(* IEC 61131-3 sources: PLC-Static-Analysis/modules/plc-rules/src/test/resources/dev/plca/rules/RulesFuzzTestInputs/fuzzRules, 23 files *)

(* ---- PLCA-Q007_compliant.st ---- *)
FUNCTION F_Twice : INT
VAR_INPUT
    n : INT;
END_VAR
F_Twice := F_Plus(n, n);
END_FUNCTION

FUNCTION F_Plus : INT
VAR_INPUT
    a : INT;
    b : INT;
END_VAR
F_Plus := a + b;
END_FUNCTION

(* ---- PLCA-P001_compliant.st ---- *)
VAR_GLOBAL
    gMode : INT;
    gOk : BOOL;
END_VAR

FUNCTION_BLOCK FB_Ok
VAR_INPUT
    bA : BOOL;
    bB : BOOL;
END_VAR
VAR_OUTPUT
    bOut : BOOL;
    nOut : INT;
END_VAR
VAR
    n : INT;
END_VAR
// default, then override in an IF
bOut := FALSE;
IF bA THEN
    bOut := TRUE;
END_IF
// latches
bOut S= bA;
bOut R= bB;
// sequential use: read in between
nOut := 1;
n := nOut * 2;
nOut := n;
// locals are not coils by default
n := 0;
n := 5;
// mutually exclusive branches
IF bA THEN
    gOk := TRUE;
ELSE
    gOk := FALSE;
END_IF
END_FUNCTION_BLOCK

PROGRAM P_Ok
VAR
    fb : FB_Ok;
END_VAR
gMode := 1;
fb(bA := gMode > 0);
gMode := 2;
END_PROGRAM

VAR_GLOBAL
    gnCycles : DINT;
END_VAR

PROGRAM P_Count
gnCycles := gnCycles + 1;
END_PROGRAM

PROGRAM P_ResetCount
gnCycles := 0;
END_PROGRAM

(* ---- PLCA-P001_locals_locals.st ---- *)
FUNCTION_BLOCK FB_L
VAR
    n : INT;
END_VAR
n := 1;
n := 2; // PLCA-P001
END_FUNCTION_BLOCK

FUNCTION F_L : INT
VAR
    n : INT;
END_VAR
n := 1;
n := 2;
F_L := n;
END_FUNCTION

(* ---- PLCA-P001_noncompliant.st ---- *)
VAR_GLOBAL
    gLamp : BOOL;
    gValve : BOOL;
END_VAR

PROGRAM P_A
VAR
    qMotor AT %QX0.0 : BOOL;
    b1 : BOOL;
    b2 : BOOL;
    tmr : TON;
END_VAR
qMotor := b1;
qMotor := b2; // PLCA-P001
gLamp := b1;
tmr(IN := b1, PT := T#1S, Q => gValve);
END_PROGRAM

PROGRAM P_B
VAR
    b : BOOL;
END_VAR
gLamp := b; // PLCA-P001
gValve := NOT b; // PLCA-P001
END_PROGRAM

FUNCTION_BLOCK FB_Out
VAR_INPUT
    bIn : BOOL;
END_VAR
VAR_OUTPUT
    bOut : BOOL;
END_VAR
bOut := bIn;
bOut := NOT bIn; // PLCA-P001
END_FUNCTION_BLOCK

(* ---- PLCA-Q001_compliant.st ---- *)
FUNCTION_BLOCK FB_Used
VAR
    nCount : INT;
    nForChildren : INT;
    aBuf : ARRAY[0..cMax] OF INT;
    nSpare1 : INT;
    bReserve_2 : BOOL;
    {attribute 'OPC.UA.DA' := '1'}
    rExposed : REAL;
    iSensor AT %I* : BOOL;
    pTarget : POINTER TO INT;
    nAddr : INT;
    nReadFromOutside : INT;
END_VAR
VAR CONSTANT
    cMax : INT := 9;
END_VAR
pTarget := ADR(nAddr);
aBuf[0] := 1;

METHOD Inc
nCount := nCount + 1;
END_METHOD
END_FUNCTION_BLOCK

FUNCTION_BLOCK FB_Child EXTENDS FB_Used
nForChildren := 0;
END_FUNCTION_BLOCK

FUNCTION_BLOCK ABSTRACT FB_Abstract_Base
VAR
    nForImplementations : INT;
END_VAR
END_FUNCTION_BLOCK

PROGRAM P_User
VAR
    fb : FB_Used;
    n : INT;
END_VAR
fb.Inc();
n := fb.nReadFromOutside;
END_PROGRAM

(* ---- PLCA-Q001_noncompliant.st ---- *)
FUNCTION_BLOCK FB_Unused
VAR_INPUT
    bIn : BOOL;
END_VAR
VAR
    nNeverUsed : INT; // PLCA-Q001
    bUsed : BOOL;
    rTemp, rOther : REAL; // PLCA-Q001 PLCA-Q001
END_VAR
VAR_TEMP
    nScratch : DINT; // PLCA-Q001
END_VAR
bUsed := bIn;
END_FUNCTION_BLOCK

PROGRAM P_Main
VAR
    fbUnused : FB_Unused;
    fbNotCalled : FB_Unused; // PLCA-Q001
    n : INT;
END_VAR
fbUnused(bIn := n > 0);
END_PROGRAM

FUNCTION F_Unused : INT
VAR_INPUT
    nIn : INT;
END_VAR
VAR
    nLocal : INT; // PLCA-Q001
END_VAR
F_Unused := nIn;
END_FUNCTION

(* ---- PLCA-Q003_compliant.st ---- *)
FUNCTION_BLOCK FB_FloatOk
VAR_INPUT
    r : REAL;
    n : INT;
END_VAR
VAR_OUTPUT
    b : BOOL;
END_VAR
VAR CONSTANT
    cA : REAL := 1.0;
    cB : REAL := 2.0;
END_VAR
b := ABS(r - 1.5) < 0.001;
b := n = 3;
b := r > 1.0;
b := cA = cB;
END_FUNCTION_BLOCK

(* ---- PLCA-Q003_noncompliant.st ---- *)
FUNCTION_BLOCK FB_Float
VAR_INPUT
    r : REAL;
    lr : LREAL;
    n : INT;
END_VAR
VAR_OUTPUT
    b : BOOL;
END_VAR
b := r = 1.5; // PLCA-Q003
IF lr <> r THEN // PLCA-Q003
    b := FALSE;
END_IF
b := n = 0.0; // PLCA-Q003
b := r * 2.0 = INT_TO_REAL(n); // PLCA-Q003
END_FUNCTION_BLOCK

(* ---- PLCA-Q004_compliant.st ---- *)
FUNCTION_BLOCK FB_DivOk
VAR_INPUT
    a : DINT;
    r : REAL;
END_VAR
VAR_OUTPUT
    q : DINT;
    rq : REAL;
END_VAR
VAR CONSTANT
    cTwo : DINT := 2;
END_VAR
q := a / cTwo;
IF a <> 0 THEN
    q := 100 / a;
END_IF
rq := r / 2.0;
q := DIV(a, cTwo);
END_FUNCTION_BLOCK

(* ---- PLCA-Q004_noncompliant.st ---- *)
FUNCTION_BLOCK FB_Div
VAR_INPUT
    a : DINT;
    r : REAL;
END_VAR
VAR_OUTPUT
    q : DINT;
    rq : REAL;
END_VAR
VAR CONSTANT
    cZero : DINT := 0;
    cTwo : DINT := 2;
END_VAR
q := a / 0; // PLCA-Q004
q := a MOD cZero; // PLCA-Q004
rq := r / 0.0; // PLCA-Q004
q := DIV(a, cTwo - 2); // PLCA-Q004
END_FUNCTION_BLOCK

(* ---- PLCA-Q005_compliant.st ---- *)
FUNCTION_BLOCK FB_LoopOk
VAR
    i : INT;
    j : INT;
    a : ARRAY[0..9] OF INT;
END_VAR
FOR i := 0 TO 9 DO
    a[i] := i;
    j := i * 2;
    FOR j := 0 TO 1 DO
        a[j] := 0;
    END_FOR
END_FOR
i := 0;
END_FUNCTION_BLOCK

(* ---- PLCA-Q005_noncompliant.st ---- *)
FUNCTION F_Inc : BOOL
VAR_IN_OUT
    nVal : INT;
END_VAR
nVal := nVal + 1;
END_FUNCTION

FUNCTION_BLOCK FB_Loop
VAR
    i : INT;
    a : ARRAY[0..9] OF INT;
END_VAR
FOR i := 0 TO 9 DO
    IF a[i] = 0 THEN
        i := i + 1; // PLCA-Q005
    END_IF
    FOR i := 0 TO 2 DO // PLCA-Q005
        a[i] := 0;
    END_FOR
    F_Inc(nVal := i); // PLCA-Q005
END_FOR
END_FUNCTION_BLOCK

(* ---- PLCA-Q006_compliant.st ---- *)
FUNCTION_BLOCK FB_InOk
VAR_INPUT
    bIn : BOOL;
    pIn : POINTER TO INT;
    refIn : REFERENCE TO INT;
END_VAR
VAR_IN_OUT
    nInOut : INT;
END_VAR
VAR
    bCopy : BOOL;
END_VAR
bCopy := bIn;
pIn^ := 1;
refIn := 2;
nInOut := 3;
END_FUNCTION_BLOCK

PROGRAM P_Caller
VAR
    fb : FB_InOk;
    n : INT;
END_VAR
fb.bIn := TRUE;
fb(bIn := FALSE, nInOut := n);
END_PROGRAM

(* ---- PLCA-Q006_noncompliant.st ---- *)
TYPE ST_Pt :
STRUCT
    x : INT;
    y : INT;
END_STRUCT
END_TYPE

FUNCTION_BLOCK FB_In
VAR_INPUT
    bIn : BOOL;
    nIn : INT;
    stIn : ST_Pt;
END_VAR
bIn := FALSE; // PLCA-Q006
stIn.x := 0; // PLCA-Q006

METHOD M
VAR_INPUT
    nArg : INT;
END_VAR
nIn := 5; // PLCA-Q006
nArg := 0; // PLCA-Q006
END_METHOD
END_FUNCTION_BLOCK

FUNCTION_BLOCK FB_In2 EXTENDS FB_In
nIn := 1; // PLCA-Q006
END_FUNCTION_BLOCK

FUNCTION F_In : INT
VAR_INPUT
    n : INT;
END_VAR
n := n + 1; // PLCA-Q006
F_In := n;
END_FUNCTION

(* ---- PLCA-Q007_noncompliant.st ---- *)
FUNCTION F_Rec : INT
VAR_INPUT
    n : INT;
END_VAR
IF n > 0 THEN
    F_Rec := F_Rec(n - 1); // PLCA-Q007
END_IF
END_FUNCTION

FUNCTION F_A : INT
VAR_INPUT
    n : INT;
END_VAR
F_A := F_B(n); // PLCA-Q007
END_FUNCTION

FUNCTION F_B : INT
VAR_INPUT
    n : INT;
END_VAR
F_B := F_A(n);
END_FUNCTION

FUNCTION_BLOCK FB_Tree
METHOD Visit : BOOL
Visit := THIS^.Visit(); // PLCA-Q007
END_METHOD
END_FUNCTION_BLOCK

(* ---- PLCA-S001_compliant.st ---- *)
FUNCTION_BLOCK FB_ConnOk
VAR_INPUT
    sPassword : STRING;
    sExpected : STRING;
END_VAR
VAR
    sPwd : STRING;
    sHost : STRING;
    sMask : STRING;
    sAms : STRING;
    sMsg : STRING;
    sVersion : STRING;
    nPasswordLength : INT;
    bOk : BOOL;
END_VAR
sPwd := '';
sHost := '127.0.0.1';
sMask := '255.255.255.0';
sAms := '5.12.34.56.1.1';
sMsg := 'Password wrong';
sVersion := '1.2.3';
sHost := '0.0.0.0';
nPasswordLength := 8;
bOk := sPassword = sExpected;
END_FUNCTION_BLOCK

(* ---- PLCA-S001_noncompliant.st ---- *)
VAR_GLOBAL
    gsPlcIp : STRING := '10.0.0.15'; // PLCA-S001
    gsApiToken : STRING := 'abc123xyz'; // PLCA-S001
END_VAR

FUNCTION_BLOCK FB_Conn
VAR_INPUT
    sPassword : STRING;
END_VAR
VAR
    sPwd : STRING;
    sHost : STRING;
    bOk : BOOL;
    fbClient : FB_TcpClient;
    wsKennwort : WSTRING := "geheim"; // PLCA-S001
END_VAR
sPwd := 'hunter2'; // PLCA-S001
sHost := '192.168.1.100:502'; // PLCA-S001
bOk := sPassword = 'letmein'; // PLCA-S001
fbClient(sRemoteHost := '172.16.0.2', sPassword := 'admin'); // PLCA-S001 PLCA-S001
END_FUNCTION_BLOCK

(* ---- PLCA-P002_compliant.st ---- *)
PROGRAM P_IoOk
VAR
    iButton AT %IX0.0 : BOOL;
    qLamp AT %QX0.1 : BOOL;
    iTemp AT %I* : INT;
END_VAR
qLamp := iButton AND iTemp > 0;
END_PROGRAM

(* ---- PLCA-P002_noncompliant.st ---- *)
PROGRAM P_Io
VAR
    b : BOOL;
    w : WORD;
END_VAR
b := %IX0.0; // PLCA-P002
%QX0.1 := b; // PLCA-P002
w := %MW10 + %IW2; // PLCA-P002 PLCA-P002
END_PROGRAM

(* ---- PLCA-Q001_globals_globals.st ---- *)
VAR_GLOBAL
    gUsed : INT;
    gNotReferenced : INT; // PLCA-Q001
    gSpareWord : WORD;
    gInit : INT := cStart;
END_VAR
VAR_GLOBAL CONSTANT
    cStart : INT := 3;
END_VAR

PROGRAM P
gUsed := gInit;
END_PROGRAM

(* ---- PLCA-Q002_compliant.st ---- *)
TYPE E_Mode : (Manual, Auto := 5, Service); END_TYPE

PROGRAM P_CaseOk
VAR
    n : INT;
    m : INT;
    eMode : E_Mode;
END_VAR
CASE n OF
    1: m := 1;
ELSE
    m := 0;
END_CASE
CASE eMode OF
    E_Mode.Manual: m := 0;
    Auto, Service: m := 1;
END_CASE
END_PROGRAM

(* ---- PLCA-Q002_noncompliant.st ---- *)
TYPE E_State : (Idle, Run, Stop); END_TYPE

PROGRAM P_Case
VAR
    n : INT;
    m : INT;
    eState : E_State;
END_VAR
CASE n OF // PLCA-Q002
    1: m := 1;
END_CASE
CASE eState OF // PLCA-Q002
    Idle: m := 0;
    Run: m := 1;
END_CASE
IF m > 0 THEN
    CASE m OF 1..5: n := 0; END_CASE // PLCA-Q002
END_IF
END_PROGRAM

(* ---- PLCA-Q002_strict_strict.st ---- *)
TYPE E_Light : (Red, Green); END_TYPE

PROGRAM P_Strict
VAR
    eLight : E_Light;
    b : BOOL;
END_VAR
CASE eLight OF // PLCA-Q002
    Red: b := FALSE;
    Green: b := TRUE;
END_CASE
END_PROGRAM
